// TIA Portal V20 export
VAR_GLOBAL   // PLC tag table "POS3.0"
   "IO-OUT-POS3_0_Regelventil_Ausgleichszylinder_Sollwert" AT %QW204 : Int;   // IO-OUT +Feld-940RN1 Regelventil Ausgleichszylinder Sollwert in mbar (IO-Link)
   "IN-POS3_0-1012B1 Kraftsensor" AT %ID4 : DWord;   // DE +Pos=3.0-1012B1 Kraftsensor
   "IO-OUT-POS3_0_Regelventil_Überlastzylinder_Sollwert" AT %QW206 : Int;   // IO-OUT +Feld-940RN2 Regelventil Überlastzylinder Sollwert in mbar (IO-Link)
   DE_POS3_0_Endlage_Überlastzylinder AT %I201.6 : Bool;   // DE+Pos=3.0-1031B3 Endlage Überlastzylinder
   "IO-IN-POS3_0_Regelventil_Ausgleichszylinder_Istwert" AT %IW204 : Int;   // IO-IN +Feld-940RN1 Regelventil Ausgleichszylinder Istwert in mbar (IO-Link)
   "IO-IN-POS3_0_Regelventil_Überlastzylinder_Istwert" AT %IW206 : Int;   // IO-IN +Feld-940RN2 Regelventil Überlastzylinder Istwert in mbar (IO-Link)
   AZ_1001T1_Pos3_0__Fixed_Out AT %I482.0 : "AZ_FixedIO_Drv2PLC";
   AZ_1001T1_Pos3_0__St_Monitor AT %I484.0 : "AZ_FixedMonitor";
   AZ_1001T1_Pos3_0__Prm_Status AT %I508.0 : "AZ_PrmRW_Drv2PLC";
   AZ_1002T1_Pos3_0_Drehachse__Fixed_Out AT %I582.0 : "AZ_FixedIO_Drv2PLC";
   AZ_1002T1_Pos3_0_Drehachse__St_Monitor AT %I584.0 : "AZ_FixedMonitor";
   AZ_1002T1_Pos3_0_Drehachse__Prm_Status AT %I608.0 : "AZ_PrmRW_Drv2PLC";
   AZ_1002T1_Pos3_0_Drehachse_AssignableMonitor AT %ID618 : DWord;
   AZ_1002T1_Pos3_0_Drehachse_AssignableMonitor1 AT %ID622 : DWord;
   AZ_1002T1_Pos3_0_Drehachse_AssignableMonitor2 AT %ID626 : DWord;
   AZ_1002T1_Pos3_0_Drehachse_AssignableMonitor3 AT %ID630 : DWord;
   AZ_1001T1_Pos3_0__OpeDataSel AT %QW498 : Word;
   AZ_1001T1_Pos3_0__Fixed_In AT %Q500.0 : "AZ_FixedIO_PLC2Drv";
   AZ_1001T1_Pos3_0__DDO AT %Q502.0 : "AZ_DDO_PLC2Drv";
   AZ_1001T1_Pos3_0__Prm_Set AT %Q526.0 : "AZ_PrmRW_PLC2Drv";
   AZ_1002T1_Pos3_0_Drehachse__OpeDataSel AT %QW598 : Word;
   AZ_1002T1_Pos3_0_Drehachse__Fixed_In AT %Q600.0 : "AZ_FixedIO_PLC2Drv";
   AZ_1002T1_Pos3_0_Drehachse__DDO AT %Q602.0 : "AZ_DDO_PLC2Drv";
   AZ_1002T1_Pos3_0_Drehachse__Prm_Set AT %Q626.0 : "AZ_PrmRW_PLC2Drv";
   "IO-IN-POS3_0_Wegmessung_Ausgleichszylinder_Istwert" AT %IW208 : Int;   // IO-IN +POS=3.0-1011B1 Wegmessung Ausgleichszylinder Istwert in mm (IO-Link)
   AZ_1002T1_Pos3_0_Drehachse__Remote_IN AT %Q596.0 : "AZ_RemoteIO_Plc2Drv";
   AZ_1001T1_Pos3_0__Remote_IN AT %Q496.0 : "AZ_RemoteIO_Plc2Drv";
   AZ_1001T1_Pos3_0__Remote_Out AT %I478.0 : "AZ_RemoteIO_Drv2Plc";
   AZ_1002T1_Pos3_0_Drehachse__Remote_Out AT %I578.0 : "AZ_RemoteIO_Drv2Plc";
END_VAR
